DATA_BLOCK "GDB_OperationsResultTest"
{ S7_Optimized_Access := 'TRUE' }
VERSION : 0.1
NON_RETAIN
VAR
    Status {ExternalWritable := 'False'} : "FRK_TestStatus";
END_VAR
BEGIN
END_DATA_BLOCK
